SUBAPPLICATION Uebung_148_AX (* Übung zu DlPgnRequest: Software Identification vom VT anfordern und empfangen *)
  (* Standard: 61499-2; Description: Copyright (c) 2026 Meisterschulen am Ostbahnhof This program and the accompanying materials are made available under the terms of the Eclipse Public License 2.0 which is available at https://www.eclipse.org/legal/epl-2.0/ SPDX-License-Identifier: EPL-2.0 *)
  (* Version 1.0, 2026-11-17, Franz Höpfinger, Meisterschulen am Ostbahnhof, initial API and implementation and/or initial documentation *)
  PACKAGE Uebungen;
  IMPORT isobus::pgn::ISO_CAN_NODE::NODE1;
  IMPORT isobus::pgn::ISOUSERHOME_e::network;
  IMPORT Uebungen::const::Uebung_120_129::Filter::VT_ADD;
  IMPORT Uebungen::const::Uebung_120_129::Filter::VT_FLT;
  IMPORT isobus::pgn::const::PgnDef::PGN_SOFTWARE_IDENTIFICATION;
  IMPORT logiBUS::io::DI::logiBUS_DI::Input_I1;
  IMPORT logiBUS::io::DI::logiBUS_DI_Events::BUTTON_SINGLE_CLICK;
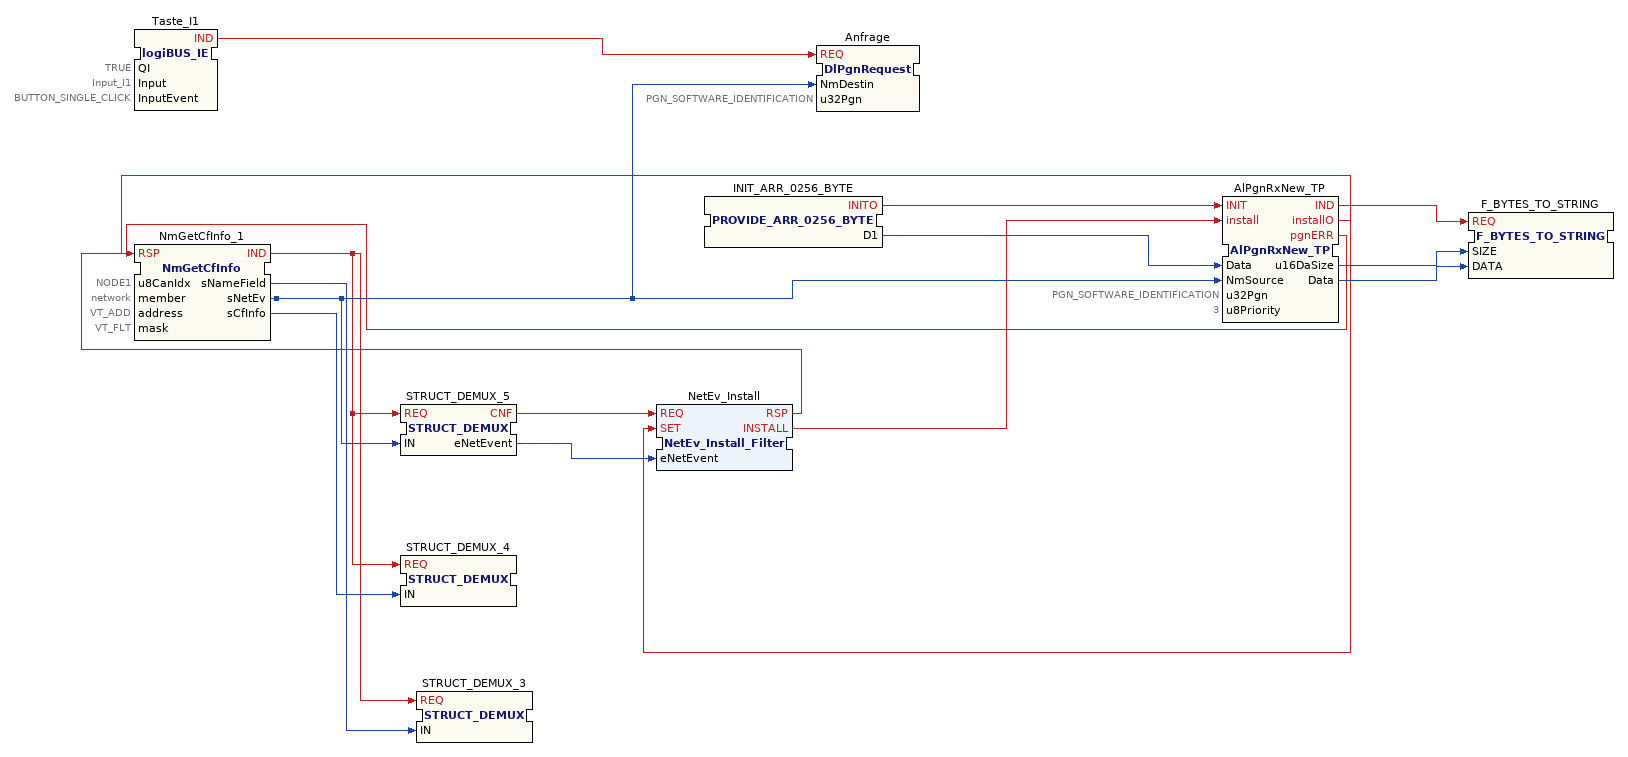
  (* DlPgnRequest: Software Identification (PGN 0xFEDA) vom VT anfordern NmGetCfInfo (network, VT-Filter) meldet den VT, AlPgnRxNew_TP wird auf 0xFEDA von ihm installiert. I1 Klick: Anfrage.REQ schickt den Request an den VT (NmDestin = sNetEv), s16Status 0 = OK. Antwort (meist TP, Felder mit * getrennt) im Watch: u16DaSize und F_BYTES_TO_STRING. *)
  FBS
    STRUCT_DEMUX_3 : eclipse4diac::convert::STRUCT_DEMUX; {SET_ATTRIBUTE(StructuredType, isobus::pgn::NAMEFIELD_T)}
    NmGetCfInfo_1 : isobus::pgn::NmGetCfInfo(u8CanIdx := NODE1, member := network, address := VT_ADD, mask := VT_FLT);
    STRUCT_DEMUX_4 : eclipse4diac::convert::STRUCT_DEMUX; {SET_ATTRIBUTE(StructuredType, isobus::pgn::CF_INFO_T)}
    STRUCT_DEMUX_5 : eclipse4diac::convert::STRUCT_DEMUX; {SET_ATTRIBUTE(StructuredType, isobus::pgn::ISONETEVENT_T)}
    INIT_ARR_0256_BYTE : eclipse4diac::convert::providers::PROVIDE_ARR_0256_BYTE;
    AlPgnRxNew_TP : isobus::pgn::rx::AlPgnRxNew_TP(u32Pgn := PGN_SOFTWARE_IDENTIFICATION, u8Priority := 3);
    F_BYTES_TO_STRING : logiBUS::utils::dyn_arr::F_BYTES_TO_STRING;
    Taste_I1 : logiBUS::io::DI::logiBUS_IE(QI := TRUE, Input := Input_I1, InputEvent := BUTTON_SINGLE_CLICK);
    Anfrage : isobus::pgn::tx::DlPgnRequest(u32Pgn := PGN_SOFTWARE_IDENTIFICATION); (* Request (PGN 0xEA00) an den VT *)
  END_FBS
  SUBAPPS
    NetEv_Install : MyLib::sys::NetEv_Install_Filter;
  END_SUBAPPS
  EVENT_CONNECTIONS
    NmGetCfInfo_1.IND TO STRUCT_DEMUX_3.REQ;
    NmGetCfInfo_1.IND TO STRUCT_DEMUX_4.REQ;
    NmGetCfInfo_1.IND TO STRUCT_DEMUX_5.REQ;
    INIT_ARR_0256_BYTE.INITO TO AlPgnRxNew_TP.INIT;
    AlPgnRxNew_TP.IND TO F_BYTES_TO_STRING.REQ;
    AlPgnRxNew_TP.installO TO NmGetCfInfo_1.RSP;
    AlPgnRxNew_TP.pgnERR TO NmGetCfInfo_1.RSP;
    STRUCT_DEMUX_5.CNF TO NetEv_Install.REQ;
    NetEv_Install.RSP TO NmGetCfInfo_1.RSP;
    AlPgnRxNew_TP.installO TO NetEv_Install.SET;
    NetEv_Install.INSTALL TO AlPgnRxNew_TP.install;
    Taste_I1.IND TO Anfrage.REQ;
  END_CONNECTIONS
  DATA_CONNECTIONS
    NmGetCfInfo_1.sNameField TO STRUCT_DEMUX_3.IN;
    NmGetCfInfo_1.sNetEv TO STRUCT_DEMUX_5.IN;
    NmGetCfInfo_1.sCfInfo TO STRUCT_DEMUX_4.IN;
    INIT_ARR_0256_BYTE.D1 TO AlPgnRxNew_TP.Data;
    AlPgnRxNew_TP.u16DaSize TO F_BYTES_TO_STRING.SIZE;
    AlPgnRxNew_TP.Data TO F_BYTES_TO_STRING.DATA;
    STRUCT_DEMUX_5.eNetEvent TO NetEv_Install.eNetEvent;
    NmGetCfInfo_1.sNetEv TO AlPgnRxNew_TP.NmSource;
    NmGetCfInfo_1.sNetEv TO Anfrage.NmDestin;
  END_CONNECTIONS
END_SUBAPPLICATION
